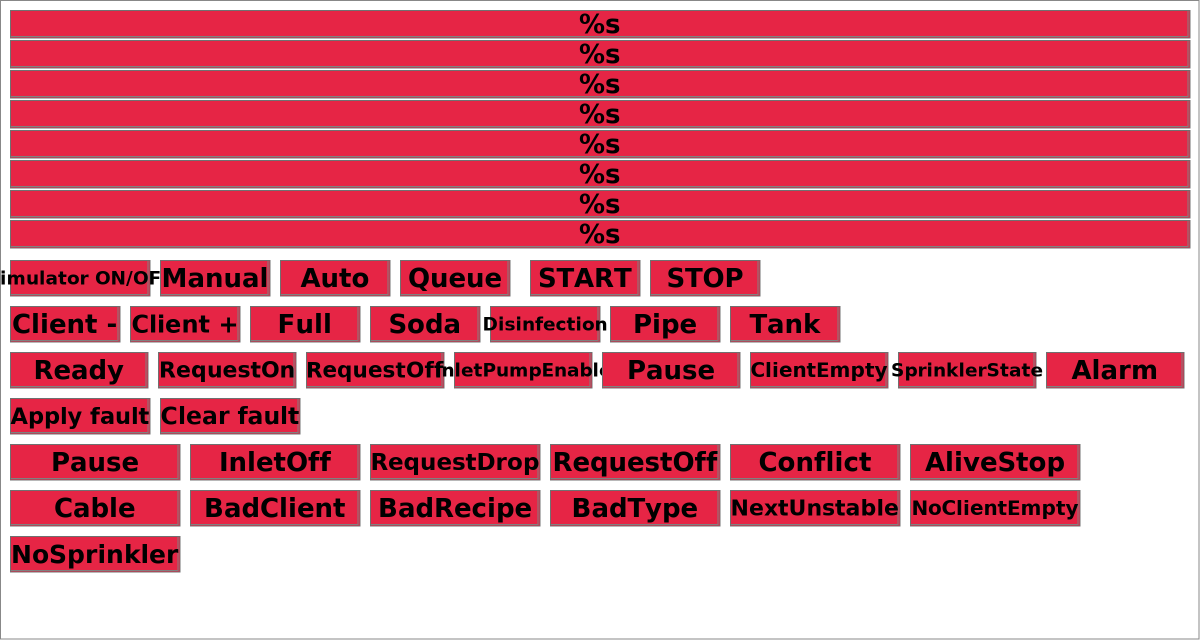
VISUALIZATION vis_SiemensSim  // 1200x640
    Button (10,10 1180x28), "%s", text variable: g_Anybus.fbSim.sSim
    Button (10,40 1180x28), "%s", text variable: g_Anybus.fbSim.sMode
    Button (10,70 1180x28), "%s", text variable: g_Anybus.fbSim.sClient
    Button (10,100 1180x28), "%s", text variable: g_Anybus.fbSim.sFault
    Button (10,130 1180x28), "%s", text variable: g_Anybus.fbSim.sFromCip
    Button (10,160 1180x28), "%s", text variable: g_Anybus.fbSim.sToCip
    Button (10,190 1180x28), "%s", text variable: g_Anybus.fbSim.sManual
    Button (10,220 1180x28), "%s", text variable: g_Anybus.fbSim.sInterface
    Button (10,260 140x36), "Simulator ON/OFF"
        OnMouseClick: execute { g_Anybus.bSimEnable:=NOT g_Anybus.bSimEnable; }
    Button (160,260 110x36), "Manual"
        OnMouseClick: execute { g_Anybus.fbSim.eMode:=E_Sim_Mode.eManual; }
    Button (280,260 110x36), "Auto"
        OnMouseClick: execute { g_Anybus.fbSim.eMode:=E_Sim_Mode.eAuto; }
    Button (400,260 110x36), "Queue"
        OnMouseClick: execute { g_Anybus.fbSim.eMode:=E_Sim_Mode.eQueue; }
    Button (530,260 110x36), "START"
        OnMouseClick: execute { g_Anybus.fbSim.bStart:=TRUE; }
    Button (650,260 110x36), "STOP"
        OnMouseClick: execute { g_Anybus.fbSim.bStop:=TRUE; }
    Button (10,306 110x36), "Client -"
        OnMouseClick: execute { IF g_Anybus.fbSim.stClient.nClient>1 THEN g_Anybus.fbSim.stClient.nClient:=g_Anybus.fbSim.stClient.nClient-1; END_IF }
    Button (130,306 110x36), "Client +"
        OnMouseClick: execute { IF g_Anybus.fbSim.stClient.nClient<30 THEN g_Anybus.fbSim.stClient.nClient:=g_Anybus.fbSim.stClient.nClient+1; END_IF }
    Button (250,306 110x36), "Full"
        OnMouseClick: execute { g_Anybus.fbSim.stClient.eRecipe:=E_Anybus_RecipeType.eFull; }
    Button (370,306 110x36), "Soda"
        OnMouseClick: execute { g_Anybus.fbSim.stClient.eRecipe:=E_Anybus_RecipeType.eDetergent; }
    Button (490,306 110x36), "Disinfection"
        OnMouseClick: execute { g_Anybus.fbSim.stClient.eRecipe:=E_Anybus_RecipeType.eDisinfectionOnly; }
    Button (610,306 110x36), "Pipe"
        OnMouseClick: execute { g_Anybus.fbSim.stClient.eType:=E_Anybus_ClientType.ePipe; }
    Button (730,306 110x36), "Tank"
        OnMouseClick: execute { g_Anybus.fbSim.stClient.eType:=E_Anybus_ClientType.eTank; }
    Button (10,352 138x36), "Ready"
        OnMouseClick: execute { g_Anybus.fbSim.stManual.bReady:=NOT g_Anybus.fbSim.stManual.bReady; }
    Button (158,352 138x36), "RequestOn"
        OnMouseClick: execute { g_Anybus.fbSim.stManual.bRequestOn:=NOT g_Anybus.fbSim.stManual.bRequestOn; }
    Button (306,352 138x36), "RequestOff"
        OnMouseClick: execute { g_Anybus.fbSim.stManual.bRequestOff:=NOT g_Anybus.fbSim.stManual.bRequestOff; }
    Button (454,352 138x36), "InletPumpEnable"
        OnMouseClick: execute { g_Anybus.fbSim.stManual.bInletPumpEnable:=NOT g_Anybus.fbSim.stManual.bInletPumpEnable; }
    Button (602,352 138x36), "Pause"
        OnMouseClick: execute { g_Anybus.fbSim.stManual.bPause:=NOT g_Anybus.fbSim.stManual.bPause; }
    Button (750,352 138x36), "ClientEmpty"
        OnMouseClick: execute { g_Anybus.fbSim.stManual.bClientEmpty:=NOT g_Anybus.fbSim.stManual.bClientEmpty; }
    Button (898,352 138x36), "SprinklerState"
        OnMouseClick: execute { g_Anybus.fbSim.stManual.bSprinklerState:=NOT g_Anybus.fbSim.stManual.bSprinklerState; }
    Button (1046,352 138x36), "Alarm"
        OnMouseClick: execute { g_Anybus.fbSim.stManual.bAlarm:=NOT g_Anybus.fbSim.stManual.bAlarm; }
    Button (10,398 140x36), "Apply fault"
        OnMouseClick: execute { g_Anybus.fbSim.bFaultOn:=TRUE; }
    Button (160,398 140x36), "Clear fault"
        OnMouseClick: execute { g_Anybus.fbSim.bFaultOn:=FALSE; }
    Button (10,444 170x36), "Pause"
        OnMouseClick: execute { g_Anybus.fbSim.eFault:=E_Sim_Fault.ePause; }
    Button (190,444 170x36), "InletOff"
        OnMouseClick: execute { g_Anybus.fbSim.eFault:=E_Sim_Fault.eInletOff; }
    Button (370,444 170x36), "RequestDrop"
        OnMouseClick: execute { g_Anybus.fbSim.eFault:=E_Sim_Fault.eRequestDrop; }
    Button (550,444 170x36), "RequestOff"
        OnMouseClick: execute { g_Anybus.fbSim.eFault:=E_Sim_Fault.eRequestOff; }
    Button (730,444 170x36), "Conflict"
        OnMouseClick: execute { g_Anybus.fbSim.eFault:=E_Sim_Fault.eConflict; }
    Button (910,444 170x36), "AliveStop"
        OnMouseClick: execute { g_Anybus.fbSim.eFault:=E_Sim_Fault.eAliveStop; }
    Button (10,490 170x36), "Cable"
        OnMouseClick: execute { g_Anybus.fbSim.eFault:=E_Sim_Fault.eCable; }
    Button (190,490 170x36), "BadClient"
        OnMouseClick: execute { g_Anybus.fbSim.eFault:=E_Sim_Fault.eBadClient; }
    Button (370,490 170x36), "BadRecipe"
        OnMouseClick: execute { g_Anybus.fbSim.eFault:=E_Sim_Fault.eBadRecipe; }
    Button (550,490 170x36), "BadType"
        OnMouseClick: execute { g_Anybus.fbSim.eFault:=E_Sim_Fault.eBadType; }
    Button (730,490 170x36), "NextUnstable"
        OnMouseClick: execute { g_Anybus.fbSim.eFault:=E_Sim_Fault.eNextUnstable; }
    Button (910,490 170x36), "NoClientEmpty"
        OnMouseClick: execute { g_Anybus.fbSim.eFault:=E_Sim_Fault.eNoClientEmpty; }
    Button (10,536 170x36), "NoSprinkler"
        OnMouseClick: execute { g_Anybus.fbSim.eFault:=E_Sim_Fault.eNoSprinkler; }
END_VISUALIZATION

(* stored: Version 1.1.0.1, ProductVersion 3.1.4026.20
   Visu vis_SiemensSim: Id {cab46f44-5473-4414-ab4d-973c938892d3} *)
